Fanuc KAREL source: kt00017.KL

-- PROVISIONAL review KL for V770-1; original PC SHA256 1704a085c8ec27d05aa116c40f7cd8792013970da5ecc62616646dec5e339401
-- Incomplete behavior may be omitted. Consult companion uncertainty JSON. Do not deploy.
PROGRAM KT00017
%NOLOCKGROUP
VAR
  I2 : INTEGER
  OUT : INTEGER
-- UNRESOLVED_DECL Y1 type=002018
BEGIN
  -- UNRESOLVED_PC offsets 5-19; opcodes 2E,22,9D,33,B2
  -- UNRESOLVED_PC offsets 24-35; opcodes 2E,23
  -- UNRESOLVED_PC offsets 40-62; opcodes 22,9D,33,B1,21,52,23
  -- UNRESOLVED_PC offsets 67-71; opcodes 7F
END KT00017
